SUBAPPLICATION Uebung_265_AX (* Dimmer mit Taster: I1 tippen = ein/aus, I1 lange druecken = stufenlos dimmen (Richtung wechselt bei jedem langen Druck), I2 = ein, I3 = aus; LED an Q1 mit logiBUS_QD_DIMMER_G (Gamma 2.2) *)
  (* Standard: 61499-2; Description: Copyright (c) 2026 Meisterschulen am Ostbahnhof This program and the accompanying materials are made available under the terms of the Eclipse Public License 2.0 which is available at https://www.eclipse.org/legal/epl-2.0/ SPDX-License-Identifier: EPL-2.0 *)
  (* Version 1.0, 2026-11-07, Franz Höpfinger, Meisterschulen am Ostbahnhof, initial API and implementation and/or initial documentation *)
  PACKAGE Uebungen;
  IMPORT logiBUS::io::DI::logiBUS_DI::Input_I1;
  IMPORT logiBUS::io::DI::logiBUS_DI::Input_I2;
  IMPORT logiBUS::io::DI::logiBUS_DI::Input_I3;
  IMPORT logiBUS::io::DI::logiBUS_DI_Events::BUTTON_LONG_PRESS_START;
  IMPORT logiBUS::io::DI::logiBUS_DI_Events::BUTTON_LONG_PRESS_UP;
  IMPORT logiBUS::io::DI::logiBUS_DI_Events::BUTTON_SINGLE_CLICK;
  IMPORT logiBUS::io::DQ::logiBUS_DO::Output_Q1;
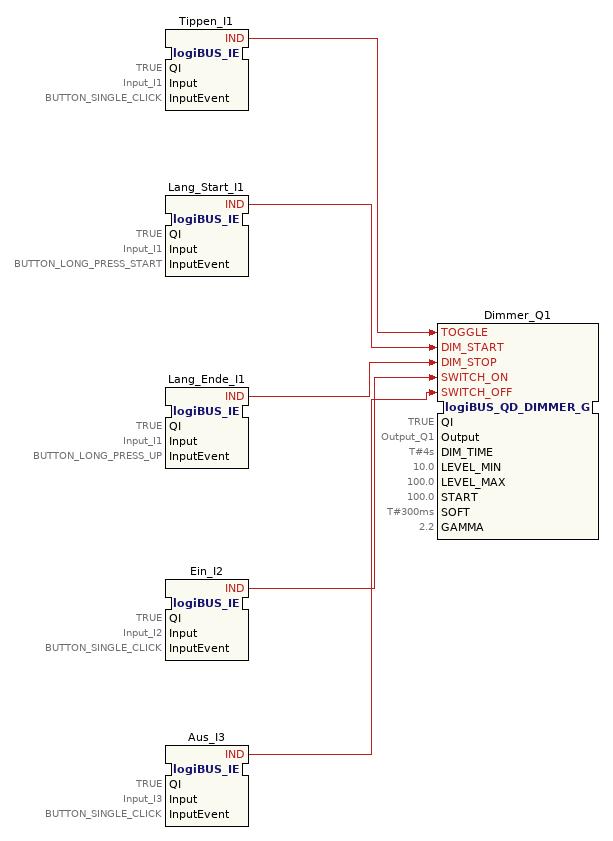
  FBS
    Tippen_I1 : logiBUS::io::DI::logiBUS_IE(QI := TRUE, Input := Input_I1, InputEvent := BUTTON_SINGLE_CLICK);
    Lang_Start_I1 : logiBUS::io::DI::logiBUS_IE(QI := TRUE, Input := Input_I1, InputEvent := BUTTON_LONG_PRESS_START);
    Lang_Ende_I1 : logiBUS::io::DI::logiBUS_IE(QI := TRUE, Input := Input_I1, InputEvent := BUTTON_LONG_PRESS_UP);
    Ein_I2 : logiBUS::io::DI::logiBUS_IE(QI := TRUE, Input := Input_I2, InputEvent := BUTTON_SINGLE_CLICK);
    Aus_I3 : logiBUS::io::DI::logiBUS_IE(QI := TRUE, Input := Input_I3, InputEvent := BUTTON_SINGLE_CLICK);
    Dimmer_Q1 : logiBUS::io::DQ::logiBUS_QD_DIMMER_G(QI := TRUE, Output := Output_Q1, DIM_TIME := T#4s, LEVEL_MIN := 10.0, LEVEL_MAX := 100.0, START := 100.0, SOFT := T#300ms, GAMMA := 2.2);
  END_FBS
  EVENT_CONNECTIONS
    Tippen_I1.IND TO Dimmer_Q1.TOGGLE;
    Lang_Start_I1.IND TO Dimmer_Q1.DIM_START;
    Lang_Ende_I1.IND TO Dimmer_Q1.DIM_STOP;
    Ein_I2.IND TO Dimmer_Q1.SWITCH_ON;
    Aus_I3.IND TO Dimmer_Q1.SWITCH_OFF;
  END_CONNECTIONS
END_SUBAPPLICATION
